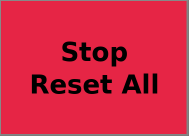
VISUALIZATION OperationButton_Stop  // 189x136
VAR_IN_OUT
	stOperation	:ST_OperationButtons;
END_VAR
    Button (0,0 189x136), "Stop Reset All", colour toggle: stOperation.bStopResetAll, pressed state: stOperation.bStopResetAll
        OnMouseClick: execute { stOperation.bStopResetAll:=TRUE; stOperation.iPauseHistory:=5; }
END_VISUALIZATION

(* stored: Version 1.1.0.1, ProductVersion 3.1.4024.13
   Visu OperationButton_Stop: Id {1e63c5c4-ebb9-43a7-be79-5a24326b4199} *)
